// TIA Portal V21 export
Screen "T12_DT"  1024x768, Number=32
  ScreenLayer 
    DateTimeField "P_DateTime" at 10,10 size 346x40
